// The ONLY place that knows the TMC event class "GenericEvents".
// Each event in that class has the text "{0}", the full text is supplied as argument.
// The class is pinned in this library (Add > Global Data Type), so it is added to the
// type system of every project that references the library.
// Used by GVL_EventDefaults.fbContext.
FUNCTION_BLOCK FB_GenericEventClass IMPLEMENTS I_EventEntryProvider
VAR
END_VAR

METHOD GetEventEntry : TcEventEntry
VAR_INPUT
	eSeverity	: TcEventSeverity;
END_VAR
CASE eSeverity OF
	TcEventSeverity.Verbose:	GetEventEntry := TC_EVENTS.GenericEvents.Verbose;
	TcEventSeverity.Info:		GetEventEntry := TC_EVENTS.GenericEvents.Info;
	TcEventSeverity.Warning:	GetEventEntry := TC_EVENTS.GenericEvents.Warning;
	TcEventSeverity.Error:		GetEventEntry := TC_EVENTS.GenericEvents.Error;
	TcEventSeverity.Critical:	GetEventEntry := TC_EVENTS.GenericEvents.Critical;
ELSE
	GetEventEntry := TC_EVENTS.GenericEvents.Error;
END_CASE
END_METHOD

END_FUNCTION_BLOCK

(* stored: Version 1.1.0.1, ProductVersion 3.1.4026.26
   POU FB_GenericEventClass: Id {1f01cc0c-e057-455b-a004-f63681b05669}, SpecialFunc None
   Method GetEventEntry: Id {5e31514b-d180-4948-8c92-03dc1d8cb51e} *)
